FUNCTION_BLOCK FIFO_UINT (* FIFO-Warteschlange fuer UINT-Werte mit frei waehlbarer Kapazitaet und Verarbeitungs-Handshake: nimmt schnelle Folgen von PUSH entgegen, liefert aber immer nur EINEN Wert per DATA aus und wartet auf PROCESSED, bevor der naechste Wert geliefert wird. *)
  (* Standard: 61499-2; Description: Copyright (c) 2026 Meisterschulen am Ostbahnhof This program and the accompanying materials are made available under the terms of the Eclipse Public License 2.0 which is available at https://www.eclipse.org/legal/epl-2.0/ SPDX-License-Identifier: EPL-2.0 *)
  (* Version 1.1, 2026-11-08, Franz Höpfinger, Meisterschulen am Ostbahnhof, RST setzt die ganze Kette zurueck (auch DELIVERING), PROCESSED wird nur bei DELIVERING angenommen, PUSH nur bei QO, QO nur bei CAPACITY > 0, CAPACITY muss aus F_LEN_ARRAY kommen. *)
  (* Version 1.0, 2026-10-13, Franz Höpfinger, Meisterschulen am Ostbahnhof, Neuentwicklung auf Basis eines alten Holobloc-FIFO_UINT-Beispiels (fixer BUF[128], DTD-Format, .serviceEvent()-Aufrufe statt echter ECC) - hier mit offenem BUF (ArraySize="*", Groesse per vorgeschalteter PROVIDE_ARR_x_UINT-Instanz + eclipse4diac::utils::arrays::F_LEN_ARRAY frei waehlbar) und echtem Request/Confirm-Verarbeitungs-Handshake auf der Konsumentenseite (DATA/PROCESSED) statt reinem Pull-on-demand. *)
  PACKAGE FIFO;
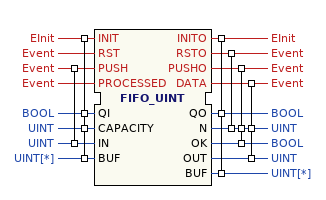
  EVENT_INPUT
    INIT : EInit WITH QI, CAPACITY, BUF; (* Service Initialization *)
    RST; (* Queue leeren und Liefer-Sperre aufheben - Reset der ganzen Kette, der Konsument muss mit zurueckgesetzt werden *)
    PUSH WITH IN; (* IN ans Ende der Queue anhaengen, falls Platz vorhanden *)
    PROCESSED; (* Konsument bestaetigt: der zuletzt per DATA gelieferte Wert ist verarbeitet. Erst danach wird (falls vorhanden) der naechste Wert per DATA geliefert. *)
  END_EVENT
  EVENT_OUTPUT
    INITO : EInit WITH QO, BUF; (* Initialisierung bestaetigt *)
    RSTO WITH N; (* Reset bestaetigt *)
    PUSHO WITH N, OK; (* PUSH bestaetigt (OK=FALSE wenn Queue voll war oder QO=FALSE) *)
    DATA WITH OUT, N; (* Ein neuer Wert ist verfuegbar. Es folgt kein weiteres DATA, bevor nicht PROCESSED eingetroffen ist. *)
  END_EVENT
  VAR_INPUT
    QI : BOOL; (* Event Input Qualifier *)
    CAPACITY : UINT; (* Kapazitaet - MUSS der Anzahl Elemente von BUF entsprechen, daher immer ueber F_LEN_ARRAY hinter der PROVIDE_ARR_x_UINT-Instanz ermitteln. Ein groesserer Wert schreibt ueber BUF hinaus. 0 ergibt QO=FALSE. *)
    IN : UINT; (* Zu pushender Wert *)
  END_VAR
  VAR_OUTPUT
    QO : BOOL; (* Event Output Qualifier *)
    N : UINT; (* Anzahl aktuell wartender (noch nicht per DATA ausgelieferter) Elemente *)
    OK : BOOL; (* TRUE wenn der letzte PUSH erfolgreich war (Queue war nicht voll und QO=TRUE) *)
    OUT : UINT; (* Zuletzt per DATA gelieferter Wert, gueltig bis zur naechsten PROCESSED-Bestaetigung *)
  END_VAR
  VAR_IN_OUT
    BUF : ARRAY [*] OF UINT; (* Ringpuffer-Speicher - Groesse wird extern ueber eine angeschlossene PROVIDE_ARR_x_UINT-Instanz vorgegeben *)
  END_VAR
  VAR
    PTR : UINT; (* Schreibposition fuer den naechsten PUSH *)
    OUTPTR : UINT; (* Leseposition fuer den naechsten auszuliefernden Wert *)
    DELIVERING : BOOL; (* TRUE = ein Wert wurde per DATA geliefert, auf PROCESSED wird gewartet *)
  END_VAR
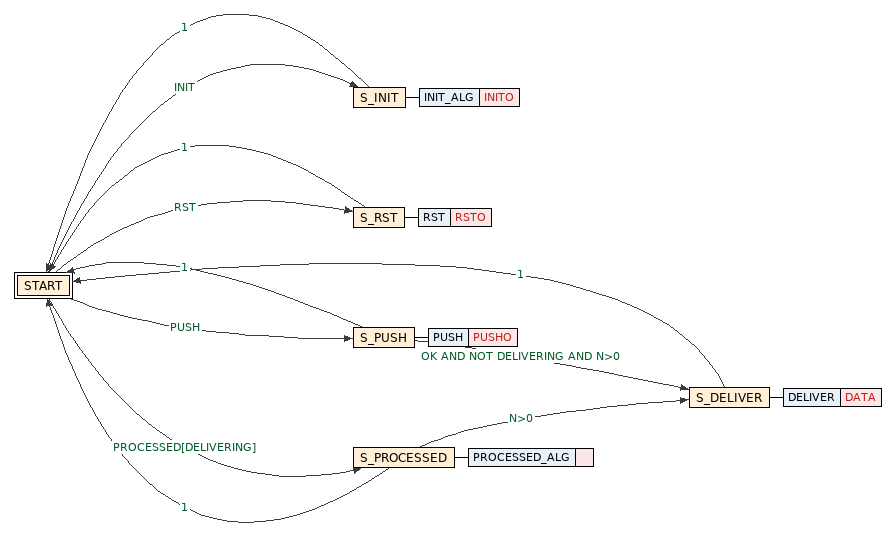
  EC_STATES
    START; (* Initial State *)
    S_INIT : INIT_ALG -> INITO;
    S_RST : RST -> RSTO;
    S_PUSH : PUSH -> PUSHO;
    S_PROCESSED : PROCESSED_ALG;
    S_DELIVER : DELIVER -> DATA; (* Naechsten Wert aus der Queue entnehmen und per DATA ausliefern *)
  END_STATES
  EC_TRANSITIONS
    START TO S_INIT := INIT;
    START TO S_RST := RST;
    START TO S_PUSH := PUSH;
    START TO S_PROCESSED := PROCESSED[DELIVERING];
    S_INIT TO START := 1;
    S_RST TO START := 1;
    S_PUSH TO S_DELIVER := OK AND NOT DELIVERING AND N>0;
    S_PUSH TO START := 1;
    S_PROCESSED TO S_DELIVER := N>0;
    S_PROCESSED TO START := 1;
    S_DELIVER TO START := 1;
  END_TRANSITIONS
  ALGORITHM INIT_ALG IN ST: (* Queue leeren und QI/QO durchreichen *)
PTR := 0;
OUTPTR := 0;
N := 0;
DELIVERING := FALSE;
OUT := 0;
OK := FALSE;
QO := QI AND CAPACITY > 0;
  END_ALGORITHM
  ALGORITHM RST IN ST: (* Queue und Liefer-Sperre leeren - RST setzt die ganze Kette zurueck, der Konsument muss mit zurueckgesetzt werden *)
PTR := 0;
OUTPTR := 0;
N := 0;
DELIVERING := FALSE;
OUT := 0;
OK := FALSE;
  END_ALGORITHM
  ALGORITHM PUSH IN ST: (* Wert anhaengen, falls Platz vorhanden *)
IF NOT QO OR N >= CAPACITY THEN
    OK := FALSE;
ELSE
    OK := TRUE;
    BUF[PTR] := IN;
    PTR := (PTR + 1) MOD CAPACITY;
    N := N + 1;
END_IF;
  END_ALGORITHM
  ALGORITHM PROCESSED_ALG IN ST: (* Liefer-Sperre aufheben - DATA fuer den naechsten Wert folgt ueber die Transition nach S_DELIVER, falls die Queue noch Elemente enthaelt *)
DELIVERING := FALSE;
  END_ALGORITHM
  ALGORITHM DELIVER IN ST: (* Vordersten Wert entnehmen und liefern *)
OUT := BUF[OUTPTR];
OUTPTR := (OUTPTR + 1) MOD CAPACITY;
N := N - 1;
DELIVERING := TRUE;
  END_ALGORITHM
END_FUNCTION_BLOCK
